(*
	FIFO queue that owns every FB_Span pointer it contains. push takes ownership and
	clears the caller's pointer; pop hands ownership back. push drops the oldest owned
	spans when the bound is reached. The bound is maxCount, but never more than
	TcOtlp_GVL.MAX_LOOP_COUNT: a maxCount of zero, or one above that limit, is held to
	MAX_LOOP_COUNT so that free always reaches the end.
	reset and next walk the spans oldest first without taking ownership. rotate moves the
	oldest span to the back, so a consumer can skip it and keep arrival order. transferTo moves the oldest spans into another queue, for handing
	a batch to an exporter.
*)
FUNCTION_BLOCK FB_SpanQueue
VAR
	_head: POINTER TO ST_LinkedListNode;
	_tail: POINTER TO ST_LinkedListNode;
	_cursor: POINTER TO ST_LinkedListNode;  // next node returned by next; 0 at the end
END_VAR
VAR_OUTPUT
	count: UDINT;
	maxCount: UDINT;
	droppedCount: UDINT;
END_VAR

(* The enforced bound: maxCount, held to MAX_LOOP_COUNT when it is zero or larger. *)
METHOD _capacity : UDINT
IF THIS^.maxCount = 0 OR THIS^.maxCount > TcOtlp_GVL.MAX_LOOP_COUNT THEN
	_capacity := TcOtlp_GVL.MAX_LOOP_COUNT;
ELSE
	_capacity := THIS^.maxCount;
END_IF
END_METHOD

METHOD FB_Exit : BOOL
VAR_INPUT
	bInCopyCode: BOOL;
END_VAR
IF NOT bInCopyCode THEN
	THIS^.free();
END_IF
END_METHOD

METHOD FB_Init : BOOL
VAR_INPUT
	bInitRetains: BOOL;
	bInCopyCode: BOOL;
	maxCount: UDINT := 0;
END_VAR
THIS^.maxCount := maxCount;
END_METHOD

(*
	Releases every owned span. push holds count to MAX_LOOP_COUNT, so the loop always
	reaches the end. If it ever stops early, the unreleased nodes stay in the queue and
	free returns FALSE, so a later call can finish the job.
*)
METHOD free : BOOL
VAR
	_idx: UDINT;
	_node: POINTER TO ST_LinkedListNode;
	_span: POINTER TO FB_Span;
END_VAR
FOR _idx := 0 TO TcOtlp_GVL.MAX_LOOP_COUNT DO
	IF THIS^._head = 0 THEN
		EXIT;
	END_IF

	_node := THIS^._head;
	THIS^._head := _node^.nxt;
	IF _node^.val <> 0 THEN
		_span := _node^.val;
		_node^.val := 0;
		_span^.delete(pSelf:=_span);
	END_IF
	__DELETE(_node);
	_node := 0;
	IF THIS^.count > 0 THEN
		THIS^.count := THIS^.count - 1;
	END_IF
END_FOR

IF THIS^._head = 0 THEN
	THIS^._tail := 0;
	THIS^.count := 0;
END_IF
THIS^._cursor := THIS^._head;
free := THIS^._head = 0;
END_METHOD

(*
	Returns the span at the cursor and advances it, or 0 after the last span. The span is
	borrowed: the queue still owns it, and it is valid only until it is popped or dropped.
	Call reset first.
*)
METHOD next : POINTER TO FB_Span
next := 0;
IF THIS^._cursor <> 0 THEN
	next := THIS^._cursor^.val;
	THIS^._cursor := THIS^._cursor^.nxt;
END_IF
END_METHOD

(* Moves the oldest span to pValue, which must be 0. The caller owns it on success. *)
METHOD pop : BOOL
VAR_IN_OUT
	pValue: POINTER TO FB_Span;
END_VAR
VAR_OUTPUT
	failureReason: E_SpanQueueFailureReason;
END_VAR
VAR
	_node: POINTER TO ST_LinkedListNode;
END_VAR
pop := FALSE;
failureReason := E_SpanQueueFailureReason.NA;

IF pValue <> 0 THEN
	failureReason := E_SpanQueueFailureReason.DESTINATION_ALREADY_ASSIGNED;
	RETURN;
END_IF
IF THIS^._head = 0 THEN
	failureReason := E_SpanQueueFailureReason.QUEUE_EMPTY;
	RETURN;
END_IF

_node := THIS^._head;
THIS^._head := _node^.nxt;
IF THIS^._head = 0 THEN
	THIS^._tail := 0;
END_IF
IF THIS^._cursor = _node THEN
	THIS^._cursor := THIS^._head;
END_IF

pValue := _node^.val;
_node^.val := 0;
_node^.nxt := 0;
__DELETE(_node);
_node := 0;
THIS^.count := THIS^.count - 1;
pop := failureReason = E_SpanQueueFailureReason.NA;
END_METHOD

(*
	Takes ownership of the span and clears pValue. On failure pValue is left unchanged
	and still owned by the caller.
*)
METHOD push : BOOL
VAR_IN_OUT
	pValue: POINTER TO FB_Span;
END_VAR
VAR_OUTPUT
	failureReason: E_SpanQueueFailureReason;
END_VAR
VAR
	_node: POINTER TO ST_LinkedListNode;
	_droppedSpan: POINTER TO FB_Span;
	_popFailureReason: E_SpanQueueFailureReason;
	_idx: UDINT;
	_bound: UDINT;
END_VAR
push := FALSE;
failureReason := E_SpanQueueFailureReason.NA;

IF pValue = 0 THEN
	failureReason := E_SpanQueueFailureReason.SPAN_POINTER_NULL;
	RETURN;
END_IF

// Allocate before evicting so an allocation failure leaves the queue unchanged.
_node := __NEW(ST_LinkedListNode);
IF _node = 0 THEN
	failureReason := E_SpanQueueFailureReason.MEMORY_ALLOCATION_FAILURE;
	RETURN;
END_IF

// maxCount is writable, so also restore the bound after a runtime reduction.
_bound := THIS^._capacity();
FOR _idx := 0 TO TcOtlp_GVL.MAX_LOOP_COUNT DO
	IF THIS^.count < _bound THEN
		EXIT;
	END_IF
	IF NOT THIS^.pop(pValue:=_droppedSpan, failureReason=>_popFailureReason) THEN
		__DELETE(_node);
		_node := 0;
		failureReason := _popFailureReason;
		RETURN;
	END_IF
	_droppedSpan^.delete(pSelf:=_droppedSpan);
	THIS^.droppedCount := THIS^.droppedCount + 1;
END_FOR
IF THIS^.count >= _bound THEN
	__DELETE(_node);
	_node := 0;
	failureReason := E_SpanQueueFailureReason.MAX_SIZE_ENFORCEMENT_FAILURE;
	RETURN;
END_IF

_node^.val := pValue;
_node^.nxt := 0;
IF THIS^._tail = 0 THEN
	THIS^._head := _node;
ELSE
	THIS^._tail^.nxt := _node;
END_IF
THIS^._tail := _node;
THIS^.count := THIS^.count + 1;
pValue := 0;
push := failureReason = E_SpanQueueFailureReason.NA;
END_METHOD

(* Moves the cursor to the oldest span, so next starts from the head. *)
METHOD reset
THIS^._cursor := THIS^._head;
END_METHOD

(*
	Moves up to count of the oldest spans into destination, which must be empty. Ownership moves
	with the nodes, so nothing is cloned or released. The move stops at this queue's count and at
	the destination's bound.
*)
METHOD transferTo : BOOL
VAR_IN_OUT
	destination: FB_SpanQueue;
END_VAR
VAR_INPUT
	count: UDINT;
END_VAR
VAR_OUTPUT
	failureReason: E_SpanQueueFailureReason;
END_VAR
VAR
	_transferCount: UDINT;
	_idx: UDINT;
END_VAR
transferTo := FALSE;
failureReason := E_SpanQueueFailureReason.NA;

IF ADR(destination) = THIS THEN
	failureReason := E_SpanQueueFailureReason.SELF_TRANSFER_NOT_ALLOWED;
	RETURN;
END_IF
IF destination.count <> 0 OR_ELSE destination._head <> 0 OR_ELSE destination._tail <> 0 THEN
	failureReason := E_SpanQueueFailureReason.DESTINATION_NOT_EMPTY;
	RETURN;
END_IF

_transferCount := MIN(count, THIS^.count, destination._capacity());
IF _transferCount = 0 THEN
	transferTo := TRUE;
	RETURN;
END_IF

// count never exceeds MAX_LOOP_COUNT, so this walk is bounded
destination._head := THIS^._head;
destination._tail := destination._head;
FOR _idx := 1 TO _transferCount - 1 DO
	destination._tail := destination._tail^.nxt;
END_FOR

THIS^._head := destination._tail^.nxt;
destination._tail^.nxt := 0;
destination._cursor := destination._head;
destination.count := _transferCount;

THIS^.count := THIS^.count - _transferCount;
THIS^._cursor := THIS^._head;
IF THIS^._head = 0 THEN
	THIS^._tail := 0;
END_IF
transferTo := TRUE;
END_METHOD

(* Moves the oldest span to the back without changing ownership, and resets the cursor. *)
METHOD rotate : BOOL
VAR_OUTPUT
	failureReason: E_SpanQueueFailureReason;
END_VAR
VAR
	_node: POINTER TO ST_LinkedListNode;
END_VAR
rotate := FALSE;
failureReason := E_SpanQueueFailureReason.NA;

IF THIS^._head = 0 THEN
	failureReason := E_SpanQueueFailureReason.QUEUE_EMPTY;
	RETURN;
END_IF

IF THIS^._head <> THIS^._tail THEN
	_node := THIS^._head;
	THIS^._head := _node^.nxt;
	_node^.nxt := 0;
	THIS^._tail^.nxt := _node;
	THIS^._tail := _node;
END_IF

THIS^._cursor := THIS^._head;
rotate := failureReason = E_SpanQueueFailureReason.NA;
END_METHOD

END_FUNCTION_BLOCK

(* stored: Version 1.1.0.1
   POU FB_SpanQueue: Id {44d433c3-56a3-4e84-9cfe-16a801713247}, SpecialFunc None
   Method _capacity: Id {2a459e68-9b56-43c7-8f56-a277c5988310}
   Method FB_Exit: Id {fd842b4a-3627-42d8-8070-91340c2c3950}
   Method FB_Init: Id {4af341fc-fbf6-4bc4-b594-12ef607990c4}
   Method free: Id {3ecf047c-8132-4a0d-bbdf-56e404d6aec4}
   Method next: Id {98c9c37a-96a9-477e-bdc0-9447f3869fa4}
   Method pop: Id {20f7cf69-8ba2-4d4e-b317-f36437396b59}
   Method push: Id {b052437c-48a1-4966-8fb6-f6eefdfa3878}
   Method reset: Id {e0e62b49-9fdc-442d-899c-23e048e89ad2}
   Method transferTo: Id {d88d0a02-dff6-4571-a522-879dc10cbe27}
   Method rotate: Id {0c8cb412-eb9c-4663-8843-2fab019dc3cb} *)
